(* PLC project Vn_op_time_to_lint, Beckhoff Automation GmbH TwinCAT PLC Control 3.5.13.21 *)
(* stored: creationDateTime 1970-01-01T00:00:00 *)

PROGRAM Vn_op_time_to_lint

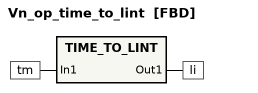
(* FBD diagram, written out as Structured Text *)
li := TIME_TO_LINT(tm);
END_PROGRAM
